{attribute 'qualified_only'}
{attribute 'strict'}
TYPE ET_AlarmType_1 : 
(
	eIdle := 0,
	eFatalError := 1,
	eError := 2,
	eWarning := 3,
	eMessage := 4,
	eHint := 5	
)INT;
END_TYPE

(* stored: Version 1.1.0.1, ProductVersion 3.1.4024.15
   DUT ET_AlarmType_1: Id {fb285c40-5606-40f8-adaf-d3a6c53c6da0} *)
